(* IEC 61131-3 sources: cps/plc, 5 files *)

(* ---- downstream.st ---- *)
PROGRAM DownstreamController
VAR
    (* Independent field sensor FC04 IR0..4 -> IW100..104. *)
    FlowRaw AT %IW100 : INT;
    WarningLimitRaw AT %IW101 : INT;
    GateObserved AT %IW102 : INT;
    SourceHealthy AT %IW103 : INT;
    SensorHeartbeat AT %IW104 : INT;
    (* PLC1 FC03 MW0..6 -> IW105..111. *)
    P1GateDesired AT %IW107 : INT;
    P1Heartbeat AT %IW111 : INT;
    (* PLC5 native FC03 MW0..13, starting address 1024. *)
    FlowSnapshot AT %MW0 : INT;
    WarningLimitSnapshot AT %MW1 : INT;
    FlowAlarmSnapshot AT %MW2 : INT;
    SensorFreshSnapshot AT %MW3 : INT;
    SensorStaleTicksSnapshot AT %MW4 : INT;
    CycleCount AT %MW5 : UINT;
    P1FreshSnapshot AT %MW6 : INT;
    P1StaleTicksSnapshot AT %MW7 : INT;
    P1DesiredSnapshot AT %MW8 : INT;
    GateObservedSnapshot AT %MW9 : INT;
    SourceHealthySnapshot AT %MW10 : INT;
    GateMismatchSnapshot AT %MW11 : INT;
    SensorHeartbeatSnapshot AT %MW12 : INT;
    P1HeartbeatSnapshot AT %MW13 : INT;
END_VAR
VAR
    SensorSeen : BOOL;
    SensorFresh : BOOL;
    P1Seen : BOOL;
    P1Fresh : BOOL;
    PreviousSensorHeartbeat : INT;
    PreviousP1Heartbeat : INT;
    SensorStaleTicks : INT;
    P1StaleTicks : INT;
    FlowAlarm : BOOL;
END_VAR

(* Each heartbeat advances independently of this controller. *)
(* Allow ~6 s for a missing heartbeat before declaring it stale. *)
IF SensorHeartbeat <> PreviousSensorHeartbeat THEN
    SensorSeen := TRUE;
    SensorStaleTicks := 0;
ELSIF SensorStaleTicks < 120 THEN
    SensorStaleTicks := SensorStaleTicks + 1;
END_IF;
PreviousSensorHeartbeat := SensorHeartbeat;
IF P1Heartbeat <> PreviousP1Heartbeat THEN
    P1Seen := TRUE;
    P1StaleTicks := 0;
ELSIF P1StaleTicks < 120 THEN
    P1StaleTicks := P1StaleTicks + 1;
END_IF;
PreviousP1Heartbeat := P1Heartbeat;
SensorFresh := SensorSeen AND (SensorStaleTicks < 120)
               AND (SourceHealthy <> 0);
P1Fresh := P1Seen AND (P1StaleTicks < 120);

(* Suppress alarms on missing upstream data, report bad quality separately. *)
FlowAlarm := SensorFresh AND (WarningLimitRaw > 0)
             AND (FlowRaw >= WarningLimitRaw);
FlowSnapshot := FlowRaw;
WarningLimitSnapshot := WarningLimitRaw;
FlowAlarmSnapshot := BOOL_TO_INT(FlowAlarm);
SensorFreshSnapshot := BOOL_TO_INT(SensorFresh);
SensorStaleTicksSnapshot := SensorStaleTicks;
P1FreshSnapshot := BOOL_TO_INT(P1Fresh);
P1StaleTicksSnapshot := P1StaleTicks;
P1DesiredSnapshot := P1GateDesired;
GateObservedSnapshot := GateObserved;
SourceHealthySnapshot := SourceHealthy;
GateMismatchSnapshot := BOOL_TO_INT(SensorFresh AND P1Fresh
                        AND (GateObserved <> P1GateDesired));
SensorHeartbeatSnapshot := SensorHeartbeat;
P1HeartbeatSnapshot := P1Heartbeat;

(* Advisory monitoring only: no outputs and no control-side writes. *)
IF CycleCount < 65535 THEN CycleCount := CycleCount + 1;
ELSE CycleCount := 0; END_IF;
END_PROGRAM

CONFIGURATION Config0
    RESOURCE Res0 ON PLC
        TASK Main(INTERVAL := T#50ms, PRIORITY := 0);
        PROGRAM Inst0 WITH Main : DownstreamController;
    END_RESOURCE
END_CONFIGURATION

(* ---- inlet.st ---- *)
PROGRAM InletController
VAR
    WaterLevelRaw AT %IW100 : INT;
    InletPosition AT %IW101 : INT;
    InletFlowRaw AT %IW102 : INT;
    InletCommand AT %QW100 : INT;
    (* Remote PLC1 %MW2..6, read through Modbus FC03 at 1026..1030. *)
    PeerGateDesired AT %IW103 : INT;
    PeerAlarm AT %IW104 : INT;
    PeerHeartbeat AT %IW107 : INT;
    LevelSnapshot AT %MW0 : INT;
    InletDesiredSnapshot AT %MW1 : INT;
    InletPositionSnapshot AT %MW2 : INT;
    InletFlowSnapshot AT %MW3 : INT;
    InletMismatchSnapshot AT %MW4 : INT;
    InletMismatchCount AT %MW5 : UINT;
    CycleCount AT %MW6 : UINT;
    PeerGateSnapshot AT %MW7 : INT;
    PeerAlarmSnapshot AT %MW8 : INT;
    PeerFreshSnapshot AT %MW9 : INT;
    PeerStaleTicksSnapshot AT %MW10 : INT;
    PeerHeartbeatSnapshot AT %MW11 : INT;
END_VAR
VAR
    WaterLevel : REAL;
    Mismatch : BOOL;
    PreviousMismatch : BOOL;
    PeerSeen : BOOL;
    PeerFresh : BOOL;
    PreviousHeartbeat : INT;
    PeerStaleTicks : INT;
END_VAR

WaterLevel := INT_TO_REAL(WaterLevelRaw) / 100.0;
IF WaterLevel > 90.0 THEN
    InletCommand := 0;
ELSIF WaterLevel > 70.0 THEN
    InletCommand := 50;
ELSE
    InletCommand := 100;
END_IF;

(* The peer scan counter changes once a second via FC03 polling. *)
(* A frozen heartbeat can indicate a stopped PLC or broken network link. *)
IF PeerHeartbeat <> PreviousHeartbeat THEN
    PeerSeen := TRUE;
    PeerStaleTicks := 0;
ELSIF PeerStaleTicks < 120 THEN
    PeerStaleTicks := PeerStaleTicks + 1;
END_IF;
PreviousHeartbeat := PeerHeartbeat;
PeerFresh := PeerSeen AND (PeerStaleTicks < 120);

(* Model-only coordination policy: if PLC1 requests a wide gate opening,
   limit inlet flow further. Missing PLC1 heartbeat closes the inlet. *)
IF NOT PeerFresh THEN
    InletCommand := 0;
ELSIF PeerAlarm <> 0 THEN
    InletCommand := 0;
ELSIF PeerGateDesired >= 75 AND InletCommand > 25 THEN
    InletCommand := 25;
END_IF;

Mismatch := InletPosition <> InletCommand;
IF Mismatch AND NOT PreviousMismatch THEN
    IF InletMismatchCount < 65535 THEN
        InletMismatchCount := InletMismatchCount + 1;
    END_IF;
END_IF;
PreviousMismatch := Mismatch;
LevelSnapshot := WaterLevelRaw;
InletDesiredSnapshot := InletCommand;
InletPositionSnapshot := InletPosition;
InletFlowSnapshot := InletFlowRaw;
InletMismatchSnapshot := BOOL_TO_INT(Mismatch);
PeerGateSnapshot := PeerGateDesired;
PeerAlarmSnapshot := PeerAlarm;
PeerFreshSnapshot := BOOL_TO_INT(PeerFresh);
PeerStaleTicksSnapshot := PeerStaleTicks;
PeerHeartbeatSnapshot := PeerHeartbeat;
IF CycleCount < 65535 THEN
    CycleCount := CycleCount + 1;
ELSE
    CycleCount := 0;
END_IF;
END_PROGRAM

CONFIGURATION Config0
    RESOURCE Res0 ON PLC
        TASK Main(INTERVAL := T#50ms, PRIORITY := 0);
        PROGRAM Inst0 WITH Main : InletController;
    END_RESOURCE
END_CONFIGURATION

(* ---- spillway.st ---- *)
PROGRAM SpillwayController
VAR
    WaterLevelRaw AT %IW100 : INT;
    GatePosition AT %IW101 : INT;
    GateCommand AT %QW100 : INT;
    (* PLC4 native FC03 MW0..3 maps to input registers 102..105. *)
    SupervisorGate AT %IW102 : INT;
    SupervisorReason AT %IW103 : INT;
    SupervisorValid AT %IW104 : INT;
    SupervisorHeartbeat AT %IW105 : INT;
    LevelSnapshot AT %MW0 : INT;
    GateSnapshot AT %MW1 : INT;
    DesiredSnapshot AT %MW2 : INT;
    AlarmSnapshot AT %MW3 : INT;
    MismatchSnapshot AT %MW4 : INT;
    MismatchCount AT %MW5 : UINT;
    CycleCount AT %MW6 : UINT;
    (* MW7..11 reserved for existing aggregate telemetry. *)
    LocalGateSnapshot AT %MW12 : INT;
    SupervisorFreshSnapshot AT %MW13 : INT;
    SupervisorGateSnapshot AT %MW14 : INT;
    SupervisorReasonSnapshot AT %MW15 : INT;
    SupervisorStaleTicksSnapshot AT %MW16 : INT;
END_VAR
VAR
    WaterLevel : REAL;
    HighLevelAlarm : BOOL;
    PreviousMismatch : BOOL;
    Mismatch : BOOL;
    LocalGate : INT;
    SupervisorSeen : BOOL;
    SupervisorFresh : BOOL;
    SupervisorPreviousHeartbeat : INT;
    SupervisorStaleTicks : INT;
END_VAR

WaterLevel := INT_TO_REAL(WaterLevelRaw) / 100.0;
HighLevelAlarm := WaterLevel > 90.0;
IF WaterLevel > 90.0 THEN
    LocalGate := 100;
ELSIF WaterLevel > 70.0 THEN
    LocalGate := 75;
ELSIF WaterLevel >= 40.0 THEN
    LocalGate := 25;
ELSE
    LocalGate := 0;
END_IF;

(* The supervisory link is optional: loss falls back to local logic. *)
IF SupervisorHeartbeat <> SupervisorPreviousHeartbeat THEN
    SupervisorSeen := TRUE;
    SupervisorStaleTicks := 0;
ELSIF SupervisorStaleTicks < 120 THEN
    SupervisorStaleTicks := SupervisorStaleTicks + 1;
END_IF;
SupervisorPreviousHeartbeat := SupervisorHeartbeat;
SupervisorFresh := SupervisorSeen AND (SupervisorStaleTicks < 120);
GateCommand := LocalGate;
(* No supervisor instruction may reduce local safety opening. *)
IF SupervisorFresh AND (SupervisorValid <> 0)
    AND (SupervisorGate > GateCommand) AND (SupervisorGate <= 100) THEN
    GateCommand := SupervisorGate;
END_IF;
LocalGateSnapshot := LocalGate;
SupervisorFreshSnapshot := BOOL_TO_INT(SupervisorFresh);
SupervisorGateSnapshot := SupervisorGate;
SupervisorReasonSnapshot := SupervisorReason;
SupervisorStaleTicksSnapshot := SupervisorStaleTicks;

Mismatch := GatePosition <> GateCommand;
IF Mismatch AND NOT PreviousMismatch THEN
    IF MismatchCount < 65535 THEN
        MismatchCount := MismatchCount + 1;
    END_IF;
END_IF;
PreviousMismatch := Mismatch;
LevelSnapshot := WaterLevelRaw;
GateSnapshot := GatePosition;
DesiredSnapshot := GateCommand;
AlarmSnapshot := BOOL_TO_INT(HighLevelAlarm);
MismatchSnapshot := BOOL_TO_INT(Mismatch);
IF CycleCount < 65535 THEN
    CycleCount := CycleCount + 1;
ELSE
    CycleCount := 0;
END_IF;
END_PROGRAM

CONFIGURATION Config0
    RESOURCE Res0 ON PLC
        TASK Main(INTERVAL := T#50ms, PRIORITY := 0);
        PROGRAM Inst0 WITH Main : SpillwayController;
    END_RESOURCE
END_CONFIGURATION

(* ---- supervisor.st ---- *)
PROGRAM SupervisoryController
VAR
    (* PLC1 FC03 MW0..12 -> local input registers 100..112. *)
    P1Level AT %IW100 : INT;
    P1GateDesired AT %IW102 : INT;
    P1HighWater AT %IW103 : INT;
    P1Heartbeat AT %IW106 : INT;
    P1LocalGate AT %IW112 : INT;
    (* PLC2 FC03 MW0..6 -> 113..119. *)
    P2InletDesired AT %IW114 : INT;
    P2Heartbeat AT %IW119 : INT;
    (* PLC3 FC03 MW0..6 -> 120..126. *)
    P3TemperatureRaw AT %IW120 : INT;
    P3TemperatureAlarm AT %IW121 : INT;
    P3GateAdvisory AT %IW122 : INT;
    P3PeerFresh AT %IW123 : INT;
    P3Heartbeat AT %IW125 : INT;
    (* Native PLC4 holding register snapshots, FC03 starting at 1024. *)
    SelectedGate AT %MW0 : INT;
    DecisionReason AT %MW1 : INT;
    DecisionValid AT %MW2 : INT;
    CycleCount AT %MW3 : UINT;
    P1FreshSnapshot AT %MW4 : INT;
    P2FreshSnapshot AT %MW5 : INT;
    P3FreshSnapshot AT %MW6 : INT;
    TemperatureAlarmSnapshot AT %MW7 : INT;
    TemperatureAdvisorySnapshot AT %MW8 : INT;
    LocalGateSnapshot AT %MW9 : INT;
    InletCommandSnapshot AT %MW10 : INT;
    HealthyPeerCount AT %MW11 : INT;
END_VAR
VAR
    P1Seen : BOOL;
    P2Seen : BOOL;
    P3Seen : BOOL;
    P1Fresh : BOOL;
    P2Fresh : BOOL;
    P3Fresh : BOOL;
    LastP1 : INT;
    LastP2 : INT;
    LastP3 : INT;
    StaleP1 : INT;
    StaleP2 : INT;
    StaleP3 : INT;
END_VAR

(* Every PLC has its own independent heartbeat; 120 scans x 50ms ~= 6s. *)
IF P1Heartbeat <> LastP1 THEN P1Seen := TRUE; StaleP1 := 0;
ELSIF StaleP1 < 120 THEN StaleP1 := StaleP1 + 1; END_IF;
IF P2Heartbeat <> LastP2 THEN P2Seen := TRUE; StaleP2 := 0;
ELSIF StaleP2 < 120 THEN StaleP2 := StaleP2 + 1; END_IF;
IF P3Heartbeat <> LastP3 THEN P3Seen := TRUE; StaleP3 := 0;
ELSIF StaleP3 < 120 THEN StaleP3 := StaleP3 + 1; END_IF;
LastP1 := P1Heartbeat;
LastP2 := P2Heartbeat;
LastP3 := P3Heartbeat;
P1Fresh := P1Seen AND (StaleP1 < 120);
P2Fresh := P2Seen AND (StaleP2 < 120);
P3Fresh := P3Seen AND (StaleP3 < 120);
P1FreshSnapshot := BOOL_TO_INT(P1Fresh);
P2FreshSnapshot := BOOL_TO_INT(P2Fresh);
P3FreshSnapshot := BOOL_TO_INT(P3Fresh);
HealthyPeerCount := BOOL_TO_INT(P1Fresh) + BOOL_TO_INT(P2Fresh) + BOOL_TO_INT(P3Fresh);
TemperatureAlarmSnapshot := P3TemperatureAlarm;
TemperatureAdvisorySnapshot := P3GateAdvisory;
LocalGateSnapshot := P1LocalGate;
InletCommandSnapshot := P2InletDesired;

(* Priority: valid high-water alarm > temperature advisory > local gate. *)
(* PLC1 remains the only gate writer. PLC4 only provides an FC03 decision. *)
DecisionValid := 0;
DecisionReason := 0;  (* 0=missing PLC1, 1=local, 2=temp, 3=high-water *)
SelectedGate := 0;
IF P1Fresh AND (P1LocalGate >= 0) AND (P1LocalGate <= 100) THEN
    DecisionValid := 1;
    SelectedGate := P1LocalGate;
    DecisionReason := 1;
    IF P1HighWater <> 0 THEN
        SelectedGate := 100;
        DecisionReason := 3;
    ELSIF P3Fresh AND (P3PeerFresh <> 0) AND (P3TemperatureAlarm <> 0)
        AND (P3GateAdvisory >= 0) AND (P3GateAdvisory <= 100)
        AND (P3GateAdvisory > SelectedGate) THEN
        SelectedGate := P3GateAdvisory;
        DecisionReason := 2;
    END_IF;
END_IF;

IF CycleCount < 65535 THEN CycleCount := CycleCount + 1;
ELSE CycleCount := 0; END_IF;
END_PROGRAM

CONFIGURATION Config0
    RESOURCE Res0 ON PLC
        TASK Main(INTERVAL := T#50ms, PRIORITY := 0);
        PROGRAM Inst0 WITH Main : SupervisoryController;
    END_RESOURCE
END_CONFIGURATION

(* ---- temperature.st ---- *)
PROGRAM TemperatureController
VAR
    (* Input registers from the independent temperature sensor, units = 0.01 C. *)
    TemperatureRaw AT %IW100 : INT;
    AlarmThresholdRaw AT %IW101 : INT;
    (* PLC1 native Modbus FC03 %MW2..6 copied into this runtime's inputs. *)
    PeerGateDesired AT %IW102 : INT;
    PeerAlarm AT %IW103 : INT;
    PeerHeartbeat AT %IW106 : INT;
    (* Read-only status and advisory, exposed on PLC3's native Modbus server. *)
    TemperatureSnapshot AT %MW0 : INT;
    TemperatureAlarmSnapshot AT %MW1 : INT;
    GateAdvisorySnapshot AT %MW2 : INT;
    PeerFreshSnapshot AT %MW3 : INT;
    PeerStaleTicksSnapshot AT %MW4 : INT;
    CycleCount AT %MW5 : UINT;
    PeerHeartbeatSnapshot AT %MW6 : INT;
END_VAR
VAR
    PeerSeen : BOOL;
    PeerFresh : BOOL;
    PreviousHeartbeat : INT;
    PeerStaleTicks : INT;
    TemperatureAlarm : BOOL;
END_VAR

(* Alarm derives from the sensor-provided temperature and threshold. *)
TemperatureAlarm := TemperatureRaw >= AlarmThresholdRaw;
TemperatureSnapshot := TemperatureRaw;
TemperatureAlarmSnapshot := BOOL_TO_INT(TemperatureAlarm);

(* Advisory ONLY. Neither PLC3 nor the HMI writes the spillway gate. *)
IF TemperatureRaw >= 3500 THEN
    GateAdvisorySnapshot := 100;
ELSIF TemperatureAlarm THEN
    GateAdvisorySnapshot := 75;
ELSE
    GateAdvisorySnapshot := 0;
END_IF;

(* PLC1 heartbeat is polled once/sec; 120 x 50 ms scans = about 6 s timeout. *)
IF PeerHeartbeat <> PreviousHeartbeat THEN
    PeerSeen := TRUE;
    PeerStaleTicks := 0;
ELSIF PeerStaleTicks < 120 THEN
    PeerStaleTicks := PeerStaleTicks + 1;
END_IF;
PreviousHeartbeat := PeerHeartbeat;
PeerFresh := PeerSeen AND (PeerStaleTicks < 120);
PeerFreshSnapshot := BOOL_TO_INT(PeerFresh);
PeerStaleTicksSnapshot := PeerStaleTicks;
PeerHeartbeatSnapshot := PeerHeartbeat;

IF CycleCount < 65535 THEN
    CycleCount := CycleCount + 1;
ELSE
    CycleCount := 0;
END_IF;
END_PROGRAM

CONFIGURATION Config0
    RESOURCE Res0 ON PLC
        TASK Main(INTERVAL := T#50ms, PRIORITY := 0);
        PROGRAM Inst0 WITH Main : TemperatureController;
    END_RESOURCE
END_CONFIGURATION
